// TIA Portal project "Clase2_PLCN3y4_variador" (V13)

(* hardware
DEVICE "S7-1200 station_1"  S7-1200 Station
   slot 0: "Rack_0"  Rack  V1.0
   slot 1: "PLC_1"  CPU 1214C AC/DC/Rly  6ES7 214-1BE30-0XB0  V2.2
*)

// ===== PLC "PLC_1"  CPU 1214C AC/DC/Rly =====

VAR_GLOBAL   // PLC tag table "Tabla de variables estándar"
   "hab" AT %I0.0 : Bool;
   "mem1" AT %M10.0 : Bool;
   "salida1" AT %Q0.0 : Bool;
   "value" AT %IW64 : UInt;
   "norm" AT %MD100 : Real;
   "scale" AT %MD120 : DWord;
   "t_conv" AT %MD200 : DWord;
   "t_out" AT %MD220 : DWord;
   "sent_giro" AT %I0.1 : Bool;
   "salida2" AT %Q0.2 : Bool;
   "Tag_1" AT %QW80 : Word;
END_VAR

// folder: System blocks/Program resources

DATA_BLOCK "TEM1"   // DB1
{ S7_Optimized_Access := 'FALSE' }
AUTHOR : Simatic
FAMILY : IEC
NAME : IEC_TMR
VERSION : 1.0
// stored: InstanceOfName ?
"?"
BEGIN
END_DATA_BLOCK

// folder: (top level)

ORGANIZATION_BLOCK "Main"   // OB1, LAD, ProgramCycle
TITLE = "Main Program Sweep (Cycle)"
{ S7_Optimized_Access := 'FALSE' }
VERSION : 0.1
// S
BEGIN

REGION Network 1
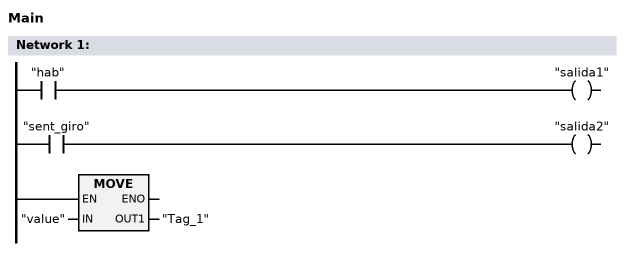
   RUNG wire#powerrail
      Contact( "hab" )
      Coil( "salida1" )
   END_RUNG
   RUNG wire#powerrail
      Contact( "sent_giro" )
      Coil( "salida2" )
   END_RUNG
   RUNG wire#powerrail
      { S7_GenerateENO := "TRUE" } Move(in := "value", out1 => "Tag_1")
   END_RUNG
   // the same network as SCL:
   "salida1" := "hab";
   "salida2" := "sent_giro";
   "Tag_1" := "value";
END_REGION
END_ORGANIZATION_BLOCK